Fanuc KAREL source: KT00486.KL

PROGRAM KT00486
%NOLOCKGROUP
VAR
  P1: POSITION
  P2: XYZWPREXT
  OUT: XYZWPREXT
BEGIN
    P2.Y = 2.0
  OUT = P1 : P2
END KT00486
